Fanuc TP program (LS listing): SpeedP.LS

/PROG  SpeedP
/ATTR
OWNER		= MNEDITOR;
COMMENT		= "RoboDK sequence";
PROG_SIZE	= 0;
CREATE		= DATE 31-12-14  TIME 12:00:00;
MODIFIED	= DATE 31-12-14  TIME 12:00:00;
FILE_NAME	= SpeedP;
VERSION		= 0;
LINE_COUNT	= 40;
MEMORY_SIZE	= 0;
PROTECT		= READ_WRITE;
TCD:  STACK_SIZE	= 0,
      TASK_PRIORITY	= 50,
      TIME_SLICE	= 0,
      BUSY_LAMP_OFF	= 0,
      ABORT_REQUEST	= 0,
      PAUSE_REQUEST	= 0;
DEFAULT_GROUP	= 1,*,*,*,*;
CONTROL_CODE	= 00000000 00000000;
/MN
   1:  ! Program generated by RoboDK v6.0.7 for Fanuc M-1iA/0.5S on XX ;
   2:  ! /XX/XXXX 18:00:00 ;
   3:  ! Using nominal kinematics. ;
   4:  PR[9,1]=1234.570 ;
   5:  PR[9,2]=-98.765 ;
   6:  PR[9,3]=50.500 ;
   7:  PR[9,4]=0.000 ;
   8:  PR[9,5]=0.000 ;
   9:  PR[9,6]=30.000 ;
  10:  UFRAME[9]=PR[9] ;
  11:  UFRAME_NUM=9 ;
  12:  PR[9,1]=10.000 ;
  13:  PR[9,2]=20.000 ;
  14:  PR[9,3]=150.000 ;
  15:  PR[9,4]=0.000 ;
  16:  PR[9,5]=0.000 ;
  17:  PR[9,6]=0.000 ;
  18:  UTOOL[9]=PR[9] ;
  19:  UTOOL_NUM=9 ;
  20:L P[1] 1mm/sec CNT0 ;
  21:J P[2] 1% CNT0 ;
  22:L P[3] 12mm/sec CNT1 ;
  23:J P[4] 3% CNT1 ;
  24:L P[5] 100mm/sec CNT2 ;
  25:J P[6] 10% CNT2 ;
  26:L P[7] 333mm/sec CNT4 ;
  27:J P[8] 22% CNT4 ;
  28:L P[9] 1000mm/sec CNT6 ;
  29:J P[10] 45% CNT6 ;
  30:L P[11] 2500mm/sec CNT9 ;
  31:J P[12] 60% CNT9 ;
  32:L P[13] 5000mm/sec CNT15 ;
  33:J P[14] 90% CNT15 ;
  34:L P[15] 12000mm/sec CNT30 ;
  35:J P[16] 100% CNT30 ;
  36:L P[17] 0mm/sec CNT75 ;
  37:J P[18] 100% CNT75 ;
  38:L P[19] 750mm/sec CNT100 ;
  39:J P[20] 1% CNT100 ;
  40:L P[21] 750mm/sec CNT100 ACC100 ;
/POS
P[1]{
   GP1:
    UF : 9, UT : 9,        CONFIG : 'L, 0, 0, 0',
	X =  -607.850  mm,	Y =   543.849  mm,	Z =   363.215  mm,
	W =  -165.000 deg,	P =    50.000 deg,	R =   150.000 deg
};
P[2]{
   GP1:
    UF : 9, UT : 9,
	J1=    10.000000 deg,	J2=    -20.000000 deg,	J3=    50.000000  mm,
	J4=    30.000000 deg
};
P[3]{
   GP1:
    UF : 9, UT : 9,        CONFIG : 'L, 0, 0, 0',
	X =  -640.584  mm,	Y =   506.980  mm,	Z =   371.534  mm,
	W =  -165.000 deg,	P =    50.000 deg,	R =   150.000 deg
};
P[4]{
   GP1:
    UF : 9, UT : 9,
	J1=    30.000000 deg,	J2=    25.000000 deg,	J3=    80.000000  mm,
	J4=    -45.000000 deg
};
P[5]{
   GP1:
    UF : 9, UT : 9,        CONFIG : 'L, 0, 0, 0',
	X =  -607.850  mm,	Y =   543.849  mm,	Z =   363.215  mm,
	W =  -165.000 deg,	P =    50.000 deg,	R =   150.000 deg
};
P[6]{
   GP1:
    UF : 9, UT : 9,
	J1=    10.000000 deg,	J2=    -20.000000 deg,	J3=    50.000000  mm,
	J4=    30.000000 deg
};
P[7]{
   GP1:
    UF : 9, UT : 9,        CONFIG : 'L, 0, 0, 0',
	X =  -640.584  mm,	Y =   506.980  mm,	Z =   371.534  mm,
	W =  -165.000 deg,	P =    50.000 deg,	R =   150.000 deg
};
P[8]{
   GP1:
    UF : 9, UT : 9,
	J1=    30.000000 deg,	J2=    25.000000 deg,	J3=    80.000000  mm,
	J4=    -45.000000 deg
};
P[9]{
   GP1:
    UF : 9, UT : 9,        CONFIG : 'L, 0, 0, 0',
	X =  -607.850  mm,	Y =   543.849  mm,	Z =   363.215  mm,
	W =  -165.000 deg,	P =    50.000 deg,	R =   150.000 deg
};
P[10]{
   GP1:
    UF : 9, UT : 9,
	J1=    10.000000 deg,	J2=    -20.000000 deg,	J3=    50.000000  mm,
	J4=    30.000000 deg
};
P[11]{
   GP1:
    UF : 9, UT : 9,        CONFIG : 'L, 0, 0, 0',
	X =  -640.584  mm,	Y =   506.980  mm,	Z =   371.534  mm,
	W =  -165.000 deg,	P =    50.000 deg,	R =   150.000 deg
};
P[12]{
   GP1:
    UF : 9, UT : 9,
	J1=    30.000000 deg,	J2=    25.000000 deg,	J3=    80.000000  mm,
	J4=    -45.000000 deg
};
P[13]{
   GP1:
    UF : 9, UT : 9,        CONFIG : 'L, 0, 0, 0',
	X =  -607.850  mm,	Y =   543.849  mm,	Z =   363.215  mm,
	W =  -165.000 deg,	P =    50.000 deg,	R =   150.000 deg
};
P[14]{
   GP1:
    UF : 9, UT : 9,
	J1=    10.000000 deg,	J2=    -20.000000 deg,	J3=    50.000000  mm,
	J4=    30.000000 deg
};
P[15]{
   GP1:
    UF : 9, UT : 9,        CONFIG : 'L, 0, 0, 0',
	X =  -640.584  mm,	Y =   506.980  mm,	Z =   371.534  mm,
	W =  -165.000 deg,	P =    50.000 deg,	R =   150.000 deg
};
P[16]{
   GP1:
    UF : 9, UT : 9,
	J1=    30.000000 deg,	J2=    25.000000 deg,	J3=    80.000000  mm,
	J4=    -45.000000 deg
};
P[17]{
   GP1:
    UF : 9, UT : 9,        CONFIG : 'L, 0, 0, 0',
	X =  -607.850  mm,	Y =   543.849  mm,	Z =   363.215  mm,
	W =  -165.000 deg,	P =    50.000 deg,	R =   150.000 deg
};
P[18]{
   GP1:
    UF : 9, UT : 9,
	J1=    10.000000 deg,	J2=    -20.000000 deg,	J3=    50.000000  mm,
	J4=    30.000000 deg
};
P[19]{
   GP1:
    UF : 9, UT : 9,        CONFIG : 'L, 0, 0, 0',
	X =  -640.584  mm,	Y =   506.980  mm,	Z =   371.534  mm,
	W =  -165.000 deg,	P =    50.000 deg,	R =   150.000 deg
};
P[20]{
   GP1:
    UF : 9, UT : 9,
	J1=    30.000000 deg,	J2=    25.000000 deg,	J3=    80.000000  mm,
	J4=    -45.000000 deg
};
P[21]{
   GP1:
    UF : 9, UT : 9,        CONFIG : 'L, 0, 0, 0',
	X =  -640.584  mm,	Y =   506.980  mm,	Z =   371.534  mm,
	W =  -165.000 deg,	P =    50.000 deg,	R =   150.000 deg
};
/END
